# EPICS autosave request: 1.5.0/debian-12/7.0.10/modules/ADCore-ee039d2/db/NDStats_settings.req
$(P)$(R)BgdWidth
$(P)$(R)ComputeStatistics
$(P)$(R)ComputeCentroid
$(P)$(R)CentroidThreshold
$(P)$(R)ComputeProfiles
$(P)$(R)CursorX
$(P)$(R)CursorY
$(P)$(R)ComputeHistogram
$(P)$(R)HistSize
$(P)$(R)HistMin
$(P)$(R)HistMax
file "NDTimeSeries_settings.req", P=$(P), R=$(R)TS:
file "NDPluginBase_settings.req", P=$(P), R=$(R)
file "sseq_settings.req", P=$(P), S=$(R)Reset
file "sseq_settings.req", P=$(P), S=$(R)Reset1
file "sseq_settings.req", P=$(P), S=$(R)Reset2
